// TwinCAT 3 PLC project Nepionic_Motion_Sandbox
// ProgramVersion: 3.1.4026.21
// libraries:
//   [Nepionic_Motion], * (Nepionic)
//   Tc2_MC2, * (Beckhoff Automation GmbH)
//   Tc3_Module, * (Beckhoff Automation GmbH)
// project tree:
//   Programs/ Main.TcPOU
//   Tasks/ PlcTask.TcTTO
// real-time tasks:
//   TASK PlcTask: cycle T#10ms, priority 20, ADS port 350
// motion (NC):
//   TASK NC-Task 1 SAF: cycle T#2ms, priority 4, ADS port 501
//   TASK NC-Task 1 SVB: cycle T#10ms, priority 8, ADS port 511
//   AXIS Axis 1 (id 1)
//     OtherSettings: AllowMotionCmdToSlave=true
//     encoder EncType=1
//     drive DrvType=5
//       Analog: TorqueSetpointScale=10, ScaleFactorActTorque=0.1
//       TimeComp: TaskDelayCycles=1
//     controller CtrType=1
//       CtrPara: PriorControlFactor=1
//         Observer: BandWidth=20
// variable links:
//   Nepionic_Motion_Sandbox/Nepionic_Motion_Sandbox Instance <-> NC-Task 1 SAF/Axes/Axis 1
//     PlcTask Inputs/Main.axis.axis_ref.NcToPlc <-> Outputs/ToPlc
//     PlcTask Outputs/Main.axis.axis_ref.PlcToNc <-> Inputs/FromPlc

CONFIGURATION Nepionic_Motion_Sandbox
    RESOURCE PLC ON TwinCAT3
        TASK PlcTask(INTERVAL := T#10ms, PRIORITY := 20);
        PROGRAM Main WITH PlcTask : Main;
    END_RESOURCE
END_CONFIGURATION

// ---- Programs/Main.TcPOU
PROGRAM Main
VAR
	axis : Mc2Axis;
	move_rel : MoveRelativeCommand(axis := axis, distance := 100, velocity := 1, acceleration := 0, deceleration := 0, jerk := 0, buffer_mode := MotionBufferMode.Aborting);
	cause_error : BOOL;
	reset_error : BOOL;
	reset_cmd : AsyncCommand;
	i : INT;
END_VAR

IF cause_error THEN
	CASE i OF
		0:
			axis.Enable();
			axis.EnablePositive();
			axis.EnableNegative();
			IF axis.IsStandstill THEN
				move_rel.Execute();
				i := 1;
			END_IF
			
		1:
			IF axis.IsConstantVelocity THEN
				axis.Disable();
				axis.DisablePositive();
				axis.DisableNegative();
				i := 2;
			END_IF
			
		2:
			IF move_rel.Error THEN
				cause_error := FALSE;
				i := 0;
			END_IF
			
	END_CASE
	
	move_rel.CyclicCall();
END_IF

IF reset_error THEN
	reset_cmd := axis.Reset();
	
	IF NOT reset_cmd.Busy THEN
		reset_error := FALSE;
	END_IF
END_IF

axis.CyclicCall();

END_PROGRAM
